FUNCTION_BLOCK PROVIDE_ARR_0008_UDINT (* FB to provide a UDINT array of size 8 (generic FB) *)
  (* Standard: 61499-2; Description: Copyright (c) 2026 Meisterschulen am Ostbahnhof This program and the accompanying materials are made available under the terms of the Eclipse Public License 2.0 which is available at https://www.eclipse.org/legal/epl-2.0/ SPDX-License-Identifier: EPL-2.0 This generic Function Block defines an array of 8 UDINT elements. Functionality: - On the INIT event, the FB reads the array 'D1' and triggers INITO. - The 'D1' InOut variable serves as the array container and can be pre-filled with initial values. - The array size can be determined with eclipse4diac::utils::arrays::F_LEN_ARRAY. Example for D1 initialization: [1, 2, ...] *)
  (* Version 1.0, 2026-11-08, Franz Höpfinger, Meisterschulen am Ostbahnhof, initial API and implementation and/or initial documentation *)
  PACKAGE eclipse4diac::convert::providers;
  {SET_ATTRIBUTE(eclipse4diac::core::GenericClassName, 'GEN_PROVIDE_ARR')}
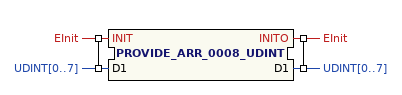
  EVENT_INPUT
    INIT : EInit WITH D1; (* Service Initialization *)
  END_EVENT
  EVENT_OUTPUT
    INITO : EInit WITH D1; (* Initialization Confirm *)
  END_EVENT
  VAR_IN_OUT
    D1 : ARRAY [0..7] OF UDINT; (* Array in/out *)
  END_VAR
END_FUNCTION_BLOCK
